// TIA Portal V21 export
TYPE "UDT_Valve"
TITLE = Задвижка
// Состояние задвижки для HMI и STL
   STRUCT
      xOpen : Bool;   // Открыта
      xClosed : Bool;   // Закрыта
      iPos_pct : Int;   // Положение, %
   END_STRUCT;
END_TYPE
